TYPE "ST_OeeSample"
VERSION : 0.1
   STRUCT
      Availability : Real;
      Performance : Real;
      Quality : Real;
      Oee : Real;
      OeeValid : Bool;
   END_STRUCT;

END_TYPE

